(* PLC project Vn_op_shr, Beckhoff Automation GmbH TwinCAT PLC Control 3.5.13.21 *)
(* stored: creationDateTime 1970-01-01T00:00:00 *)

PROGRAM Vn_op_shr

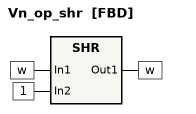
(* FBD diagram, written out as Structured Text *)
w := SHR(w, 1);
END_PROGRAM
